// TIA Portal V21 export
// export: Created 2026-11-11T00:48:15.9507755Z, ExportSetting WithDefaults, DisplayName Totally Integrated Automation Portal, DisplayVersion V21 Update 3, DisplayName STEP 7 Professional, DisplayVersion V21 Update 3, DisplayName STEP 7 Safety, DisplayVersion V21, DisplayName Tech WebApplication, DisplayVersion V21, DisplayName WinCC Basic/Comfort/Advanced, DisplayVersion V21 Update 3, DisplayName WinCC Unified, DisplayVersion V21 Update 3
FUNCTION_BLOCK "FB_Scl_sl039"   // FB60, SCL
{ S7_Optimized_Access := 'TRUE' }
VERSION : 0.1
// stored: AutoNumber true, IsIECCheckEnabled false, IsRetainMemResEnabled false, MemoryReserve 100, SetENOAutomatically false, UDAEnableTagReadback false
   VAR_INPUT
      v_src_array : Byte;
   END_VAR
   VAR_OUTPUT
      v_ret : Byte;
   END_VAR
   VAR_IN_OUT
      v_dest_variable : Variant;
      v_pos : DInt;
   END_VAR
BEGIN
   #v_ret := Deserialize(SRC_ARRAY := #v_src_array, DEST_VARIABLE => #v_dest_variable, POS := #v_pos);
END_FUNCTION_BLOCK
